(*
SPDX-FileCopyrightText: © 2026 Oleksandr Tiutyk <trofimich@gmail.com>
SPDX-License-Identifier: MIT
License: https://opensource.org/license/mit
*)

(*!
<summary>Identifies the next root scheduling or reporting action.</summary>
*)

{attribute 'qualified_only'}
{attribute 'strict'}
{attribute 'to_string'}
TYPE TEST_RUN_PHASE :
(
	STARTING,
	RUNNING_ELEMENTS,
	REPORTING_TOTALS,
	COMPLETED
);
END_TYPE

(* stored: Version 1.1.0.1
   DUT TEST_RUN_PHASE: Id {28fb3fa3-9d37-43ae-a909-28ff50ca84ca} *)
